// TIA Portal V20 export
// export: Created 2026-11-12T11:17:34.0857573Z, ExportSetting WithDefaults, DisplayName Totally Integrated Automation Portal, DisplayVersion V20, DisplayName TIA Portal Openness, DisplayVersion V20, DisplayName TIA Portal Teamcenter Gateway, DisplayVersion V20, DisplayName TIA Portal Version Control Interface, DisplayVersion V20, DisplayName STEP 7 Professional, DisplayVersion V20, DisplayName STEP 7 CFC, DisplayVersion V20, DisplayName STEP 7 Safety, DisplayVersion V20, DisplayName WinCC Basic/Comfort/Advanced, DisplayVersion V20, DisplayName SIMATIC Visualization Architect, DisplayVersion V20, DisplayName WinCC Professional, DisplayVersion V20, DisplayName SIMATIC Visualization Architect, DisplayVersion V20, DisplayName WinCC Unified, DisplayVersion V20, DisplayName SIMATIC Visualization Architect, DisplayVersion V20
TYPE "UDT_Entradas_Stopper"
// stored: IsFailsafeCompliant false
   STRUCT
      Sensor_ind_0 : Bool;   // Entrada Sensor inductivo 0 (Extremo derecho)
      Sensor_ind_1 : Bool;   // Entrada Sensor inductivo 1
      Sensor_ind_2 : Bool;   // Entrada Sensor inductivo 2
      Sensor_ind_3 : Bool;   // Entrada Sensor inductivo 3 (Extremo izquierdo)
      Reservado_E2_4 : Bool;
      Reservado_E2_5 : Bool;
      Reservado_E2_6 : Bool;
      Sensor_stopper_abajo : Bool;   // Entrada Stopper abajo
   END_STRUCT;
END_TYPE
